(* IEC 61131-3 sources: trust-platform/editors/vscode/media/examples/hmi-starter/src, 2 files *)

(* ---- config.st ---- *)
CONFIGURATION Config
RESOURCE MainRes ON PLC
    TASK MainTask (INTERVAL := T#10ms, PRIORITY := 1);
    PROGRAM Main WITH MainTask : Main;
END_RESOURCE
END_CONFIGURATION

(* ---- Main.st ---- *)
PROGRAM Main
VAR
    level   : INT;
    running : BOOL;
END_VAR
    running := TRUE;
    level := (level + 1) MOD 100;
END_PROGRAM
